// TIA Portal V21 export
// export: Created 2026-11-21T13:54:30.788407Z, ExportSetting WithDefaults, DisplayName Totally Integrated Automation Portal, DisplayVersion V21, DisplayName STEP 7 Professional, DisplayVersion V21, DisplayName STEP 7 Safety, DisplayVersion V21, DisplayName Tech WebApplication, DisplayVersion V21, DisplayName WinCC Basic/Comfort/Advanced, DisplayVersion V21, DisplayName WinCC Unified, DisplayVersion V21
VAR_GLOBAL   // PLC tag table "Pump"
   Pump_Speed AT %MW10 : Int;   // Speed of the pump
   Pump_On AT %M0.0 : Bool;   // The pump runs
   Flow AT %MD20 : Real;   // Flow through the pump
END_VAR
